Staubli VAL3: utButton.dtx

public utAppearance Appearance
  [0]
    string sBackgroundColour
    string sBackgroundImage
    string sColour
    bool bVisibility
public utBorder Border
  [0]
    string sBorderColour
public utCommon Common
  [0]
    bool bDisabled
    string sText
    string sID
    string sPage
public utText Text
  [0]
    string sFontFamily
    string sFontStyle
    string sFontWeight
    string sTextAlignment
    num nFontSize
public utEvents Events
  [0]
    bool bClick
    bool bMouseDown
    bool bMouseUp
public utData Data
  [0]
    num nVal
    bool bStatus
